// TwinCAT 3 PLC project RobotskaRokaPLC
// ProgramVersion: 3.1.4026.27
// libraries:
//   Tc2_Standard, * (Beckhoff Automation GmbH)
//   Tc2_System, * (Beckhoff Automation GmbH)
// project tree:
//   GVLs/ IO.TcGVL
//   / PlcTask.TcTTO
//   POUs/ FB_CommandSelector.TcPOU, FB_MotorControl.TcPOU, MAIN.TcPOU
// real-time tasks:
//   TASK PlcTask: cycle T#10ms, priority 20, ADS port 350
//   TASK PlcTask1: cycle T#10ms, priority 21, ADS port 351
// I/O:
//   DEVICE Device 1 (EtherCAT), AmsNetId 10.99.109.205.2.1
//     Term 1 (EK1200) [EK1200-7000 EtherCAT Power supply (1,5A E-Bus)]
//       Term 2 (EL1859) [EL1859 8Ch. Dig. Input 24V, 3ms, 8Ch. Dig. Output 24V, 0.5A]
//       Term 3 (EL1859) [EL1859 8Ch. Dig. Input 24V, 3ms, 8Ch. Dig. Output 24V, 0.5A]
//       Term 4 (EL9011) [EL9011 End Terminal]
//   DEVICE Device 2 (NOV-DP-RAM)
//   DEVICE Device 3 (CX7000), AmsNetId 10.99.109.205.4.1
//     Term 1 (CX7028) [CX7028-0000-0118]
//       modules: Module 1 (DIO_2x), Module 3 (DIO_2x), Module 5 (DI_2x), Module 7 (DI_2x)
// variable links:
//   RobotskaRokaPLC/RobotskaRokaPLC Instance <-> Device 1 (EtherCAT)/Term 1 (EK1200)/Term 2 (EL1859)
//     PlcTask Inputs/MAIN.bExtendLimit <-> Channel 3/Input
//     PlcTask Inputs/MAIN.bGripLimit <-> Channel 7/Input
//     PlcTask Inputs/MAIN.bLiftLimit <-> Channel 5/Input
//     PlcTask Inputs/MAIN.bRotateLimit <-> Channel 1/Input
//     PlcTask Outputs/MAIN.bExtendDirection <-> Channel 11/Output
//     PlcTask Outputs/MAIN.bExtendRun <-> Channel 12/Output
//     PlcTask Outputs/MAIN.bGripDirection <-> Channel 15/Output
//     PlcTask Outputs/MAIN.bGripRun <-> Channel 16/Output
//     PlcTask Outputs/MAIN.bLiftDirection <-> Channel 13/Output
//     PlcTask Outputs/MAIN.bLiftRun <-> Channel 14/Output
//     PlcTask Outputs/MAIN.bRotateDirection <-> Channel 9/Output
//     PlcTask Outputs/MAIN.bRotateRun <-> Channel 10/Output
//   RobotskaRokaPLC/RobotskaRokaPLC Instance <-> Device 3 (CX7000)/Term 1 (CX7028)
//     PlcTask Inputs/MAIN.bExtend <-> Module 5 (DI_2x)/DI_2x Input Channel 1/Input
//     PlcTask Inputs/MAIN.bManualMode <-> Module 7 (DI_2x)/DI_2x Inputs Channel 1/Input
//     PlcTask Inputs/MAIN.bRetract <-> Module 5 (DI_2x)/DI_2x Input Channel 2/Input
//     PlcTask Inputs/MAIN.bRotateLeft <-> Module 1 (DIO_2x)/DIO_2x Inputs Channel 2/Input
//     PlcTask Inputs/MAIN.bRotateRight <-> Module 3 (DIO_2x)/DIO_2x Input Channel 1/Input
//     PlcTask Inputs/MAIN.bShift <-> Module 3 (DIO_2x)/DIO_2x Input Channel 2/Input
//     PlcTask Inputs/MAIN.bStopButton <-> Module 1 (DIO_2x)/DIO_2x Inputs Channel 1/Input

CONFIGURATION RobotskaRokaPLC
    RESOURCE PLC ON TwinCAT3
        TASK PlcTask(INTERVAL := T#10ms, PRIORITY := 21);
        PROGRAM MAIN WITH PlcTask : MAIN;
    END_RESOURCE
END_CONFIGURATION

// ---- GVLs/IO.TcGVL
{attribute 'qualified_only'}
VAR_GLOBAL
	ToggleSwitch : BOOL;
    ButtonRed : BOOL;
    ButtonGreen : BOOL;

    ButtonBlackLeftUp : BOOL;
    ButtonBlackRightUp : BOOL;
    ButtonBlackLeftDown : BOOL;
    ButtonBlackRightDown : BOOL;

    SwitchReferenceRotate : BOOL;
    SwitchStepRotate : BOOL;

    SwitchReferenceExtend : BOOL;
    SwitchStepExtend : BOOL;

    SwitchReferenceLift : BOOL;
    SwitchStepLift : BOOL;

    SwitchReferenceGrip : BOOL;
    SwitchStepGrip : BOOL;
	
	LEDRed : BOOL;
    LEDGreen : BOOL;
    LEDBlueUp : BOOL;
    LEDBlueDown : BOOL;

    MotorRotateDirection : BOOL;
    MotorRotateMovement : BOOL;

    MotorExtendDirection : BOOL;
    MotorExtendMovement : BOOL;

    MotorLiftDirection : BOOL;
    MotorLiftMovement : BOOL;

    MotorGripDirection : BOOL;
    MotorGripMovement : BOOL;
END_VAR

// ---- POUs/MAIN.TcPOU
PROGRAM MAIN
VAR
    bManualMode AT %I* : BOOL;
    bRotateLeft AT %I* : BOOL;
    bRotateRight AT %I* : BOOL;
    bExtend AT %I* : BOOL;
    bRetract AT %I* : BOOL;
    bShift AT %I* : BOOL;
    bStopButton AT %I* : BOOL;

    bRotateLimit AT %I* : BOOL;
    bExtendLimit AT %I* : BOOL;
    bLiftLimit AT %I* : BOOL;
    bGripLimit AT %I* : BOOL;
	
	bAllButtonsReleased : BOOL;
	bShiftSelected : BOOL;
	bShiftMismatch : BOOL;
	bCommandArmed : BOOL;
	bMotionEnabled : BOOL;

    bRotateLeftCmd : BOOL;
    bRotateRightCmd : BOOL;
    bExtendCmd : BOOL;
    bRetractCmd : BOOL;
    bLiftUp : BOOL;
    bLiftDown : BOOL;
    bGripOpen : BOOL;
    bGripClose : BOOL;

    bReqRotateForward : BOOL;
    bReqRotateBackward : BOOL;
    bReqExtendForward : BOOL;
    bReqExtendBackward : BOOL;
    bReqLiftForward : BOOL;
    bReqLiftBackward : BOOL;
    bReqGripForward : BOOL;
    bReqGripBackward : BOOL;

    bRotateRun AT %Q* : BOOL;
    bRotateDirection AT %Q* : BOOL;

    bExtendRun AT %Q* : BOOL;
    bExtendDirection AT %Q* : BOOL;

    bLiftRun AT %Q* : BOOL;
    bLiftDirection AT %Q* : BOOL;

    bGripRun AT %Q* : BOOL;
    bGripDirection AT %Q* : BOOL;


    fbRotateSelector : FB_CommandSelector;
    fbExtendSelector : FB_CommandSelector;
    fbLiftSelector : FB_CommandSelector;
    fbGripSelector : FB_CommandSelector;

    fbRotateMotor : FB_MotorControl;
    fbExtendMotor : FB_MotorControl;
    fbLiftMotor : FB_MotorControl;
    fbGripMotor : FB_MotorControl;
	
	nSelectedMotor : INT := 0;
END_VAR

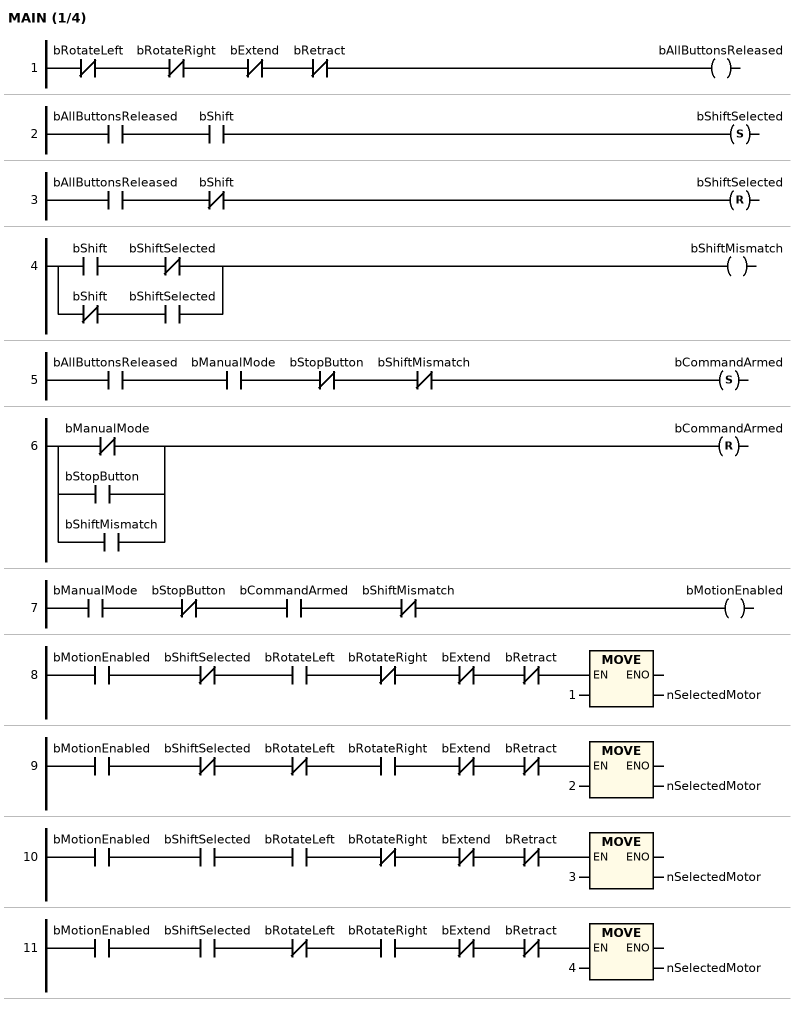
// NETWORK 1
bAllButtonsReleased := NOT bRotateLeft AND NOT bRotateRight AND NOT bExtend AND NOT bRetract;

// NETWORK 2
bShiftSelected S= bAllButtonsReleased AND bShift;

// NETWORK 3
bShiftSelected R= bAllButtonsReleased AND NOT bShift;

// NETWORK 4
bShiftMismatch := bShift AND NOT bShiftSelected OR NOT bShift AND bShiftSelected;

// NETWORK 5
bCommandArmed S= bAllButtonsReleased AND bManualMode AND NOT bStopButton AND NOT bShiftMismatch;

// NETWORK 6
bCommandArmed R= NOT bManualMode OR bStopButton OR bShiftMismatch;

// NETWORK 7
bMotionEnabled := bManualMode AND NOT bStopButton AND bCommandArmed AND NOT bShiftMismatch;

// NETWORK 8
IF bMotionEnabled AND NOT bShiftSelected AND bRotateLeft AND NOT bRotateRight AND NOT bExtend AND NOT bRetract THEN
    nSelectedMotor := 1;
END_IF

// NETWORK 9
IF bMotionEnabled AND NOT bShiftSelected AND NOT bRotateLeft AND bRotateRight AND NOT bExtend AND NOT bRetract THEN
    nSelectedMotor := 2;
END_IF

// NETWORK 10
IF bMotionEnabled AND bShiftSelected AND bRotateLeft AND NOT bRotateRight AND NOT bExtend AND NOT bRetract THEN
    nSelectedMotor := 3;
END_IF

// NETWORK 11
IF bMotionEnabled AND bShiftSelected AND NOT bRotateLeft AND bRotateRight AND NOT bExtend AND NOT bRetract THEN
    nSelectedMotor := 4;
END_IF

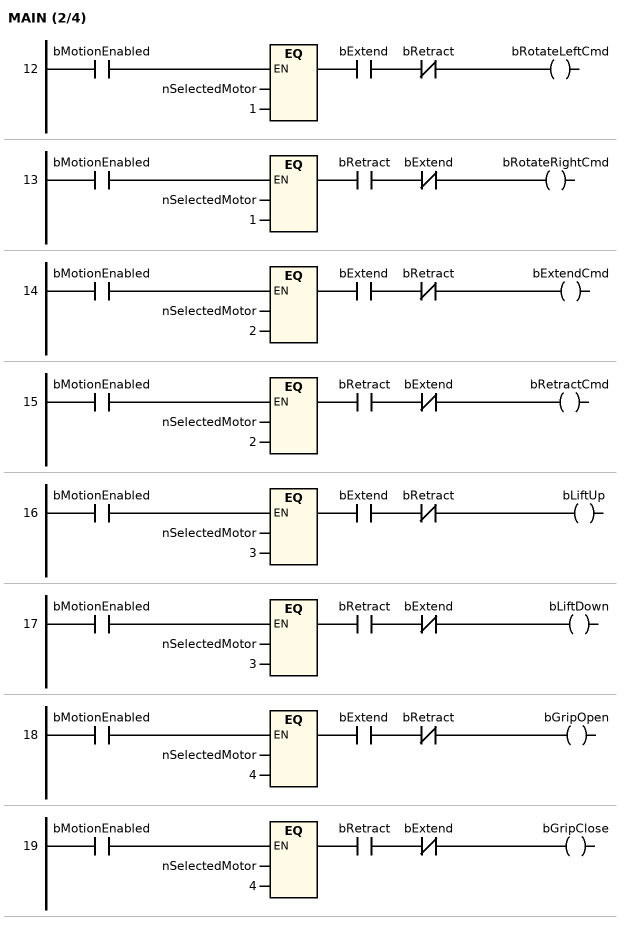
// NETWORK 12
bRotateLeftCmd := (bMotionEnabled AND nSelectedMotor = 1) AND bExtend AND NOT bRetract;

// NETWORK 13
bRotateRightCmd := (bMotionEnabled AND nSelectedMotor = 1) AND bRetract AND NOT bExtend;

// NETWORK 14
bExtendCmd := (bMotionEnabled AND nSelectedMotor = 2) AND bExtend AND NOT bRetract;

// NETWORK 15
bRetractCmd := (bMotionEnabled AND nSelectedMotor = 2) AND bRetract AND NOT bExtend;

// NETWORK 16
bLiftUp := (bMotionEnabled AND nSelectedMotor = 3) AND bExtend AND NOT bRetract;

// NETWORK 17
bLiftDown := (bMotionEnabled AND nSelectedMotor = 3) AND bRetract AND NOT bExtend;

// NETWORK 18
bGripOpen := (bMotionEnabled AND nSelectedMotor = 4) AND bExtend AND NOT bRetract;

// NETWORK 19
bGripClose := (bMotionEnabled AND nSelectedMotor = 4) AND bRetract AND NOT bExtend;

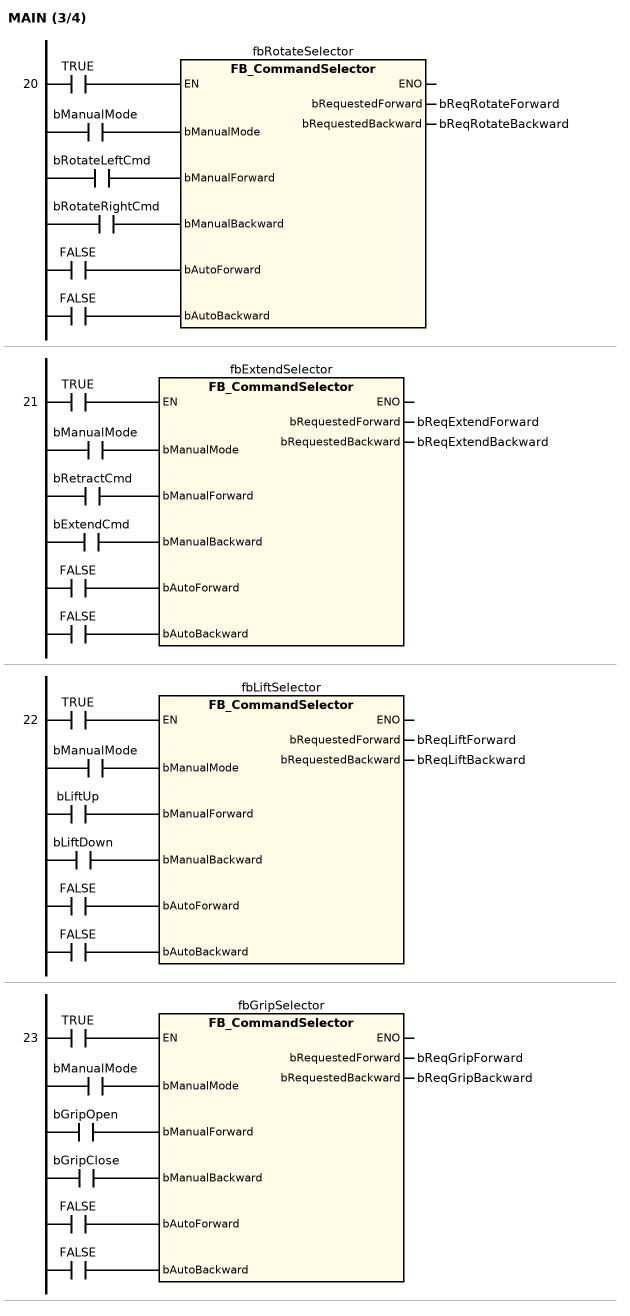
// NETWORK 20
fbRotateSelector(
    bManualMode := bManualMode,
    bManualForward := bRotateLeftCmd,
    bManualBackward := bRotateRightCmd,
    bAutoForward := FALSE,
    bAutoBackward := FALSE,
    bRequestedForward => bReqRotateForward,
    bRequestedBackward => bReqRotateBackward); // FB_CommandSelector

// NETWORK 21
fbExtendSelector(
    bManualMode := bManualMode,
    bManualForward := bRetractCmd,
    bManualBackward := bExtendCmd,
    bAutoForward := FALSE,
    bAutoBackward := FALSE,
    bRequestedForward => bReqExtendForward,
    bRequestedBackward => bReqExtendBackward); // FB_CommandSelector

// NETWORK 22
fbLiftSelector(
    bManualMode := bManualMode,
    bManualForward := bLiftUp,
    bManualBackward := bLiftDown,
    bAutoForward := FALSE,
    bAutoBackward := FALSE,
    bRequestedForward => bReqLiftForward,
    bRequestedBackward => bReqLiftBackward); // FB_CommandSelector

// NETWORK 23
fbGripSelector(
    bManualMode := bManualMode,
    bManualForward := bGripOpen,
    bManualBackward := bGripClose,
    bAutoForward := FALSE,
    bAutoBackward := FALSE,
    bRequestedForward => bReqGripForward,
    bRequestedBackward => bReqGripBackward); // FB_CommandSelector

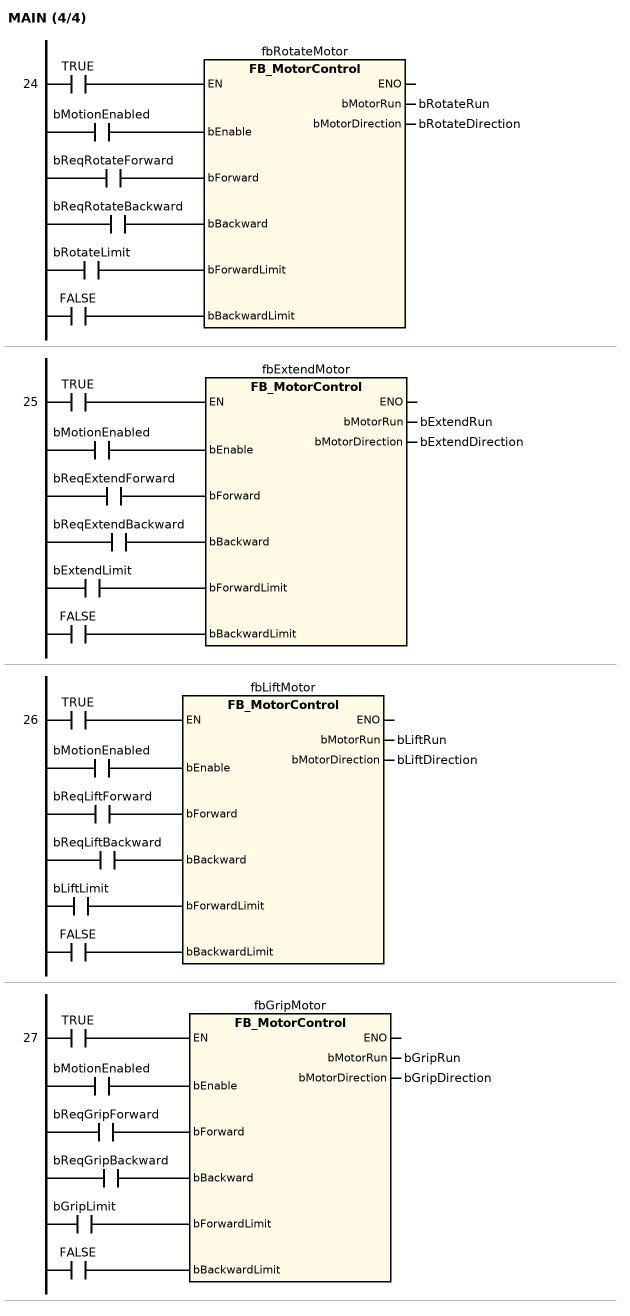
// NETWORK 24
fbRotateMotor(
    bEnable := bMotionEnabled,
    bForward := bReqRotateForward,
    bBackward := bReqRotateBackward,
    bForwardLimit := bRotateLimit,
    bBackwardLimit := FALSE,
    bMotorRun => bRotateRun,
    bMotorDirection => bRotateDirection); // FB_MotorControl

// NETWORK 25
fbExtendMotor(
    bEnable := bMotionEnabled,
    bForward := bReqExtendForward,
    bBackward := bReqExtendBackward,
    bForwardLimit := bExtendLimit,
    bBackwardLimit := FALSE,
    bMotorRun => bExtendRun,
    bMotorDirection => bExtendDirection); // FB_MotorControl

// NETWORK 26
fbLiftMotor(
    bEnable := bMotionEnabled,
    bForward := bReqLiftForward,
    bBackward := bReqLiftBackward,
    bForwardLimit := bLiftLimit,
    bBackwardLimit := FALSE,
    bMotorRun => bLiftRun,
    bMotorDirection => bLiftDirection); // FB_MotorControl

// NETWORK 27
fbGripMotor(
    bEnable := bMotionEnabled,
    bForward := bReqGripForward,
    bBackward := bReqGripBackward,
    bForwardLimit := bGripLimit,
    bBackwardLimit := FALSE,
    bMotorRun => bGripRun,
    bMotorDirection => bGripDirection); // FB_MotorControl

END_PROGRAM

// ---- POUs/FB_CommandSelector.TcPOU
FUNCTION_BLOCK FB_CommandSelector
VAR_INPUT
	bManualMode : BOOL;
    bManualForward : BOOL;
    bManualBackward : BOOL;
    bAutoForward : BOOL;
    bAutoBackward : BOOL;
END_VAR

VAR_OUTPUT
	bRequestedForward : BOOL;
    bRequestedBackward : BOOL;
END_VAR

VAR
	
END_VAR

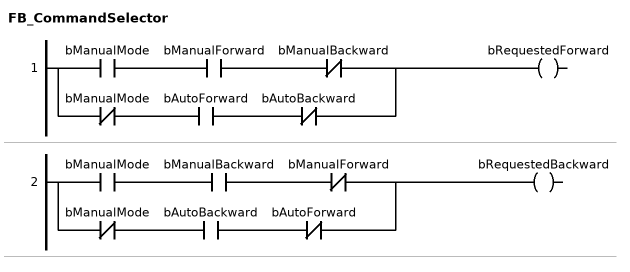
// NETWORK 1
bRequestedForward := bManualMode AND bManualForward AND NOT bManualBackward OR NOT bManualMode AND bAutoForward AND NOT bAutoBackward;

// NETWORK 2
bRequestedBackward := bManualMode AND bManualBackward AND NOT bManualForward OR NOT bManualMode AND bAutoBackward AND NOT bAutoForward;

END_FUNCTION_BLOCK

// ---- POUs/FB_MotorControl.TcPOU
FUNCTION_BLOCK FB_MotorControl
VAR_INPUT
	bEnable : BOOL;
    bForward : BOOL;
    bBackward : BOOL;
    bForwardLimit : BOOL;
    bBackwardLimit : BOOL;
END_VAR

VAR_OUTPUT
	bMotorRun : BOOL;
    bMotorDirection : BOOL;
END_VAR

VAR
	bAllowedForward : BOOL;
    bAllowedBackward : BOOL;
	bDirectionChange : BOOL;
	bDelayElapsed : BOOL;
	
	fbDirectionDelay: TON;
	tDirectionElapsed : TIME;
END_VAR

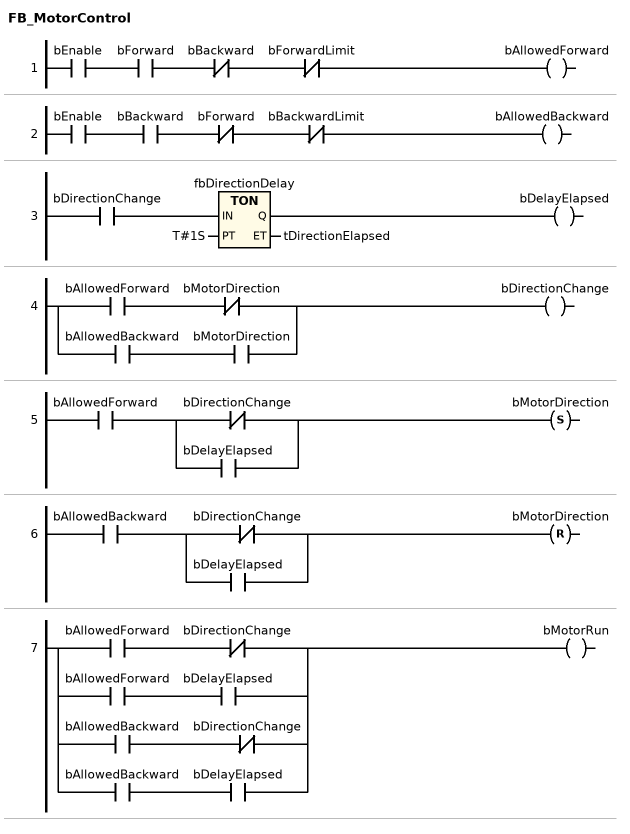
// NETWORK 1
bAllowedForward := bEnable AND bForward AND NOT bBackward AND NOT bForwardLimit;

// NETWORK 2
bAllowedBackward := bEnable AND bBackward AND NOT bForward AND NOT bBackwardLimit;

// NETWORK 3
fbDirectionDelay(IN := bDirectionChange, PT := T#1S, ET => tDirectionElapsed); // TON
bDelayElapsed := fbDirectionDelay.Q;

// NETWORK 4
bDirectionChange := bAllowedForward AND NOT bMotorDirection OR bAllowedBackward AND bMotorDirection;

// NETWORK 5
bMotorDirection S= bAllowedForward AND (NOT bDirectionChange OR bDelayElapsed);

// NETWORK 6
bMotorDirection R= bAllowedBackward AND (NOT bDirectionChange OR bDelayElapsed);

// NETWORK 7
bMotorRun := bAllowedForward AND NOT bDirectionChange OR bAllowedForward AND bDelayElapsed OR bAllowedBackward AND NOT bDirectionChange OR bAllowedBackward AND bDelayElapsed;

END_FUNCTION_BLOCK
